PROGRAM MAIN
VAR
	power1:mc_power;
	Axis1: AXIS_REF;
	jog1:mc_jog;
	moveobs:mc_moveabsolute;
	moveobs1:mc_moveabsolute;
	enable: BOOL;
	Execute: BOOL;
	JogBackwards: BOOL;
	JogForward: BOOL;
	Position: LREAL;
	Velocity: LREAL;
	Execute1: BOOL;
END_VAR

apower();
	jog1(
	Axis:=Axis1 , 
	JogForward:=JogForward, 
	JogBackwards:=JogBackwards , 
	Mode:= , 
	Position:= , 
	Velocity:= , 
	Acceleration:= , 
	Deceleration:= , 
	Jerk:= , 
	Done=> , 
	Busy=> , 
	Active=> , 
	CommandAborted=> , 
	Error=> , 
	ErrorID=> );
	moveobs(
	Axis:=Axis1 , 
	Execute:=Execute , 
	Position:= Position, 
	Velocity:=Velocity , 
	Acceleration:= , 
	Deceleration:= , 
	Jerk:= , 
	BufferMode:= , 
	Options:= , 
	Done=> , 
	Busy=> , 
	Active=> , 
	CommandAborted=> , 
	Error=> , 
	ErrorID=> );
	moveobs1(
	Axis:=Axis1 , 
	Execute:=Execute1 , 
	Position:= Position, 
	Velocity:=Velocity , 
	Acceleration:= , 
	Deceleration:= , 
	Jerk:= , 
	BufferMode:= , 
	Options:= , 
	Done=> , 
	Busy=> , 
	Active=> , 
	CommandAborted=> , 
	Error=> , 
	ErrorID=> );

ACTION apower:
power1(
	Axis:=Axis1 , 
	Enable:=enable , 
	Enable_Positive:=1 , 
	Enable_Negative:=1 , 
	Override:= , 
	BufferMode:= , 
	Options:= , 
	Status=> , 
	Busy=> , 
	Error=> , 
	ErrorID=> );
END_ACTION

END_PROGRAM

(* stored: Version 1.1.0.1, ProductVersion 3.1.4024.16
   POU MAIN: Id {84992476-be26-4e39-bd1c-ea53bae116a0}, SpecialFunc None
   Action apower: Id {0c1d298f-2ece-469f-8cc0-1a9e87f2a2c2} *)
